// TwinCAT 3 PLC project PLC
// ProgramVersion: 3.1.4026.19
// libraries:
//   Tc2_Standard, * (Beckhoff Automation GmbH)
//   Tc2_System, * (Beckhoff Automation GmbH)
//   Tc3_Vision, * (Beckhoff Automation GmbH)
// project tree:
//   / PlcTask.TcTTO
//   POUs/ MAIN.TcPOU
// real-time tasks:
//   TASK PlcTask: cycle T#10ms, priority 20, ADS port 350
//   TASK VnTask ImgAcq (Camera1): cycle T#1ms, priority 5, ADS port 351
//   TASK VnTask ADS (Camera1): cycle T#10ms, priority 6, ADS port 352
// I/O:
//   DEVICE Device 1 (RT-Ethernet Adapter)

CONFIGURATION PLC
    RESOURCE PLC ON TwinCAT3
        TASK PlcTask(INTERVAL := T#10ms, PRIORITY := 20);
        PROGRAM MAIN WITH PlcTask : MAIN;
    END_RESOURCE
END_CONFIGURATION

// ---- POUs/MAIN.TcPOU
PROGRAM MAIN
VAR
 
fbCameraControl     :    FB_VN_GevCameraControl;
eState              :    ETcVnCameraState;
hr                  :    HRESULT;

// Raw Image (Mono8 from camera)
ipImageIn           :    ITcVnImage;
ipImageInDisp       :    ITcVnDisplayableImage;

// Processed display image (RGB for colored overlays)
ipImageRGB          :    ITcVnImage;
ipImageResDisp      :    ITcVnDisplayableImage;

// QR Code
ipCodeDecodedList   :    ITcVnContainer; 
ipCodeContourList   :    ITcVnContainer;
sCodeAsString       :    STRING(255);
bCodeFound          :    BOOL := FALSE;
hrQr                :    HRESULT;
nQrAttempt          :    USINT;

// Color - RGBA format: Red
aColorRed           :    TcVnVector4_LREAL := [255, 0, 0, 255];
sDisplayText        :    STRING(512);

END_VAR

eState := fbCameraControl.GetState();

CASE eState OF
      TCVN_CS_ERROR:
        fbCameraControl.Reset();
 
      TCVN_CS_INITIAL,
      TCVN_CS_OPENING,
      TCVN_CS_OPENED,
      TCVN_CS_STARTACQUISITION:
        // Start acquisition when camera is ready.
        hr := fbCameraControl.StartAcquisition();
  
      TCVN_CS_ACQUIRING:
        // Get current Mono8 image from camera.
        hr := fbCameraControl.GetCurrentImage(ipImageIn);
  
        IF SUCCEEDED(hr) AND ipImageIn <> 0 THEN
          // Raw display image.
          hr := F_VN_CopyIntoDisplayableImage(ipImageIn, ipImageInDisp, hr);
      
          // Adaptive multi-pass QR reading.
          bCodeFound := FALSE;
          sCodeAsString := '';
          sDisplayText := '';
          ipCodeDecodedList := 0;
          ipCodeContourList := 0;

          FOR nQrAttempt := 1 TO 3 DO
            hrQr := 0;

            CASE nQrAttempt OF
              1:
                // Normal polarity and orientation.
                hrQr := F_VN_ReadQRCodeExp(
                  ipSrcImage      :=  ipImageIn,
                  ipDecodedData   :=  ipCodeDecodedList,
                  ipContours      :=  ipCodeContourList,
                  nCodeNumber     :=  1,
                  eSearchStrategy :=  TCVN_CSS_ONLY_NOT_INVERTED + TCVN_CSS_ONLY_NOT_FLIPPED,
                  hrPrev          :=  hrQr
                );
              2:
                // Allow inverted polarity.
                hrQr := F_VN_ReadQRCodeExp(
                  ipSrcImage      :=  ipImageIn,
                  ipDecodedData   :=  ipCodeDecodedList,
                  ipContours      :=  ipCodeContourList,
                  nCodeNumber     :=  1,
                  eSearchStrategy :=  TCVN_CSS_ONLY_NOT_FLIPPED,
                  hrPrev          :=  hrQr
                );
              3:
                // Allow flipped orientation.
                hrQr := F_VN_ReadQRCodeExp(
                  ipSrcImage      :=  ipImageIn,
                  ipDecodedData   :=  ipCodeDecodedList,
                  ipContours      :=  ipCodeContourList,
                  nCodeNumber     :=  1,
                  eSearchStrategy :=  TCVN_CSS_ONLY_NOT_INVERTED,
                  hrPrev          :=  hrQr
                );
            END_CASE

            IF SUCCEEDED(hrQr) AND ipCodeDecodedList <> 0 THEN
              bCodeFound := TRUE;
              hr := F_VN_ExportSubContainer_String(ipCodeDecodedList, 0, sCodeAsString, 255, hr);
              EXIT;
            END_IF
          END_FOR
          
          // Convert Mono8 to RGB for colored overlays.
          hr := F_VN_ConvertColorSpace(ipImageIn, ipImageRGB, TCVN_CST_GRAY_TO_RGB, hr);

          // Draw overlays on RGB image.
          IF bCodeFound AND ipCodeContourList <> 0 THEN
            hr := F_VN_DrawContours(ipCodeContourList, 0, ipImageRGB, aColorRed, 3, hr);
            sDisplayText := CONCAT('QR: ', sCodeAsString);
          ELSE
            sDisplayText := 'No QR Code Found';
          END_IF
          
          // Text overlay.
          hr := F_VN_PutTextExp(sDisplayText, ipImageRGB, 50, 100, ETcVnFontType.TCVN_FT_HERSHEY_SIMPLEX, 1.0, aColorRed, 2, TCVN_LT_8_CONNECTED, FALSE, hr);
          
          // Processed display image.
          hr := F_VN_CopyIntoDisplayableImage(ipImageRGB, ipImageResDisp, hr);
        END_IF
  
      TCVN_CS_STOPACQUISITION:
        ;
      TCVN_CS_TRIGGERING:
        ;
      TCVN_CS_CLOSING:
        ;  
END_CASE

END_PROGRAM
